# EPICS autosave request: examples/test/motorRecord/autosave/req/auto_positions.req
# double
$(P):Axis1.DVAL
$(P):Axis1.MFLG
